FUNCTION_BLOCK Recipe1 (* Basic Function Block Type *)
  (* Standard: 61499-2 *)
  (* Version 0.0, 10/11/2026, macie, nxtControl GmBH, Template *)
  PACKAGE Main;
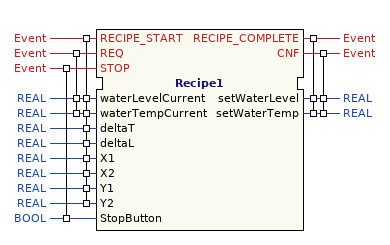
  EVENT_INPUT
    RECIPE_START WITH waterLevelCurrent, waterTempCurrent, deltaT, deltaL, X1, X2, Y1, Y2; (* Initialization Request *)
    REQ WITH waterLevelCurrent, waterTempCurrent; (* Normal Execution Request *)
    STOP WITH StopButton;
  END_EVENT
  EVENT_OUTPUT
    RECIPE_COMPLETE WITH setWaterLevel, setWaterTemp; (* Initialization Confirm *)
    CNF WITH setWaterLevel, setWaterTemp; (* Execution Confirmation *)
  END_EVENT
  VAR_INPUT
    waterLevelCurrent : REAL;
    waterTempCurrent : REAL; (* Input event qualifier *)
    deltaT : REAL;
    deltaL : REAL;
    X1 : REAL;
    X2 : REAL;
    Y1 : REAL;
    Y2 : REAL;
    StopButton : BOOL;
  END_VAR
  VAR_OUTPUT
    setWaterLevel : REAL; (* Output event qualifier *)
    setWaterTemp : REAL;
  END_VAR
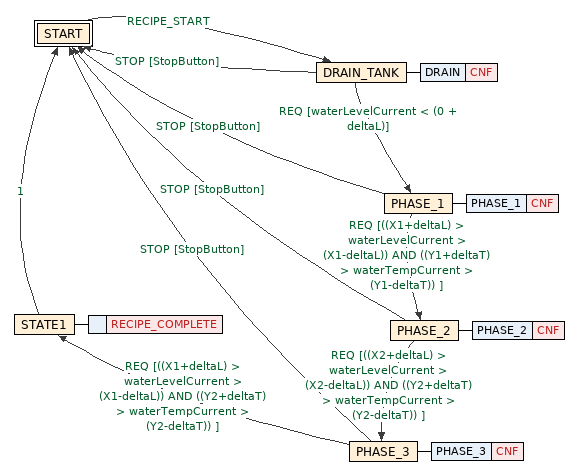
  EC_STATES
    START; (* Initial State *)
    DRAIN_TANK : DRAIN -> CNF;
    PHASE_1 : PHASE_1 -> CNF;
    PHASE_2 : PHASE_2 -> CNF;
    PHASE_3 : PHASE_3 -> CNF;
    STATE1 : -> RECIPE_COMPLETE;
  END_STATES
  EC_TRANSITIONS
    START TO DRAIN_TANK := RECIPE_START;
    DRAIN_TANK TO PHASE_1 := REQ [waterLevelCurrent < (0 + deltaL)];
    PHASE_1 TO PHASE_2 := REQ [((X1+deltaL) > waterLevelCurrent > (X1-deltaL)) AND ((Y1+deltaT) > waterTempCurrent > (Y1-deltaT)) ];
    PHASE_2 TO PHASE_3 := REQ [((X2+deltaL) > waterLevelCurrent > (X2-deltaL)) AND ((Y2+deltaT) > waterTempCurrent > (Y2-deltaT)) ];
    PHASE_3 TO STATE1 := REQ [((X1+deltaL) > waterLevelCurrent > (X1-deltaL)) AND ((Y2+deltaT) > waterTempCurrent > (Y2-deltaT)) ];
    STATE1 TO START := 1;
    DRAIN_TANK TO START := STOP [StopButton];
    PHASE_1 TO START := STOP [StopButton];
    PHASE_2 TO START := STOP [StopButton];
    PHASE_3 TO START := STOP [StopButton];
  END_TRANSITIONS
  ALGORITHM INIT IN ST: (* Initialization algorithm *)
;
  END_ALGORITHM
  ALGORITHM REQ IN ST: (* Normally executed algorithm *)
;
  END_ALGORITHM
  ALGORITHM DRAIN IN ST:
;
setWaterLevel := 0;
setWaterTemp := 0;
  END_ALGORITHM
  ALGORITHM PHASE_1 IN ST:
;
setWaterLevel := X1;
setWaterTemp := Y1;
  END_ALGORITHM
  ALGORITHM PHASE_2 IN ST:
;
setWaterLevel := X2;
setWaterTemp := Y2;
  END_ALGORITHM
  ALGORITHM PHASE_3 IN ST:
;
setWaterLevel := X1;
setWaterTemp := Y2;
  END_ALGORITHM
END_FUNCTION_BLOCK
